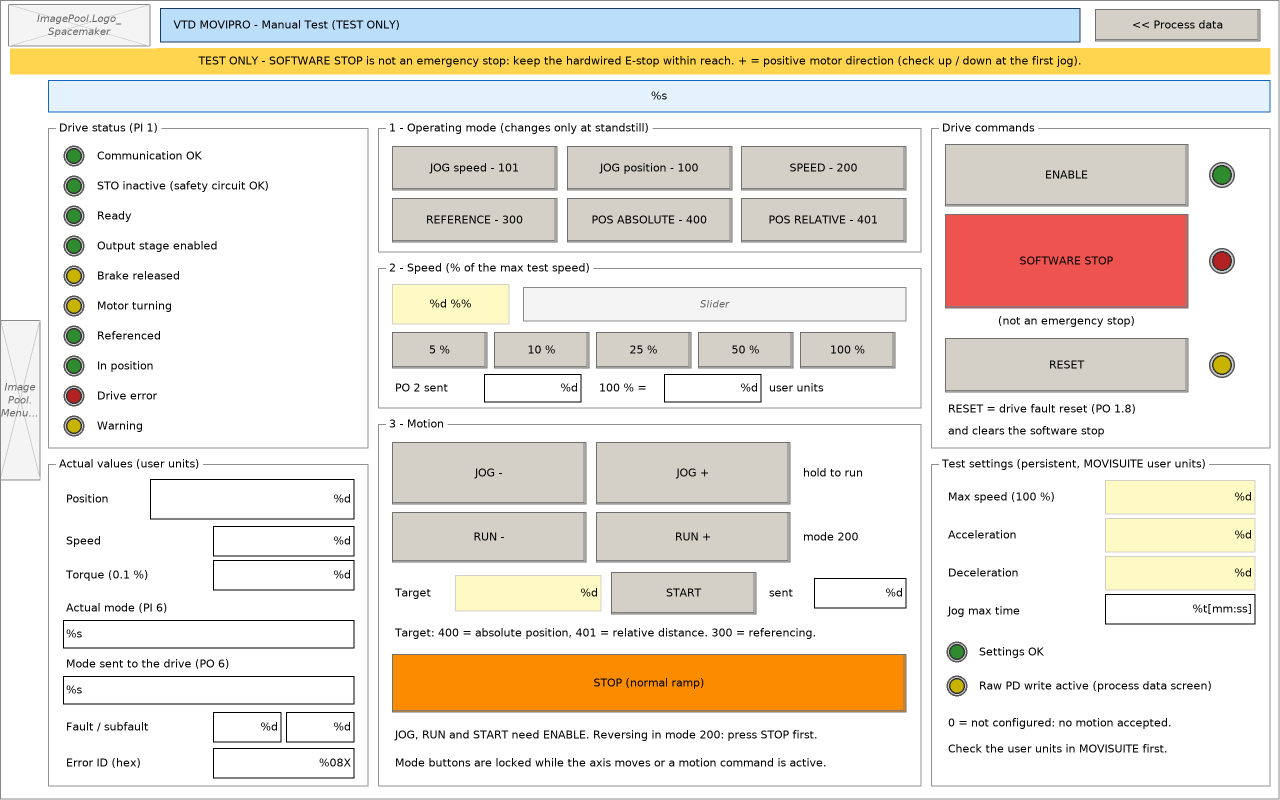
VISUALIZATION VTDManualTest  // 1280x800
    Rectangle (160,8 920x34), "VTD MOVIPRO - Manual Test (TEST ONLY)"
    Button (1095,9 165x32), "<< Process data"
        OnMouseClick: change screen: Visualization
    Rectangle (10,48 1260x26), "TEST ONLY - SOFTWARE STOP is not an emergency stop: keep the hardwired E-stop within reach. + = positive motor direction (check up / down at the first jog)."
    Rectangle (48,80 1222x32), "%s", text variable: GVL_HMI_VTD.stManualStatus.sMessage, colour toggle: GVL_HMI_VTD.stManualStatus.bMessageAlarm
    GroupBox (48,120 320x328), "Drive status (PI 1)"
    Lamp1 (62,144 24x24), variable: GVL_HMI_VTD.stManualStatus.stDrive.bCommunicationOk, style: Lamp-Lamp1-Green
    Rectangle (94,142 261x28), "Communication OK"
    Lamp1 (62,174 24x24), variable: GVL_HMI_VTD.stManualStatus.stDrive.bStoInactive, style: Lamp-Lamp1-Green
    Rectangle (94,172 261x28), "STO inactive (safety circuit OK)"
    Lamp1 (62,204 24x24), variable: GVL_HMI_VTD.stManualStatus.stDrive.bReady, style: Lamp-Lamp1-Green
    Rectangle (94,202 261x28), "Ready"
    Lamp1 (62,234 24x24), variable: GVL_HMI_VTD.stManualStatus.stDrive.bOutputStageEnabled, style: Lamp-Lamp1-Green
    Rectangle (94,232 261x28), "Output stage enabled"
    Lamp1 (62,264 24x24), variable: GVL_HMI_VTD.stManualStatus.stDrive.bBrakeReleased, style: Lamp-Lamp1-Yellow
    Rectangle (94,262 261x28), "Brake released"
    Lamp1 (62,294 24x24), variable: GVL_HMI_VTD.stManualStatus.stDrive.bMotorTurning, style: Lamp-Lamp1-Yellow
    Rectangle (94,292 261x28), "Motor turning"
    Lamp1 (62,324 24x24), variable: GVL_HMI_VTD.stManualStatus.stDrive.bReferenced, style: Lamp-Lamp1-Green
    Rectangle (94,322 261x28), "Referenced"
    Lamp1 (62,354 24x24), variable: GVL_HMI_VTD.stManualStatus.stDrive.bInPosition, style: Lamp-Lamp1-Green
    Rectangle (94,352 261x28), "In position"
    Lamp1 (62,384 24x24), variable: GVL_HMI_VTD.stManualStatus.stDrive.bError, style: Lamp-Lamp1-Red
    Rectangle (94,382 261x28), "Drive error"
    Lamp1 (62,414 24x24), variable: GVL_HMI_VTD.stManualStatus.stDrive.bWarning, style: Lamp-Lamp1-Yellow
    Rectangle (94,412 261x28), "Warning"
    GroupBox (48,456 320x330), "Actual values (user units)"
    Rectangle (63,484 82x30), "Position"
    Rectangle (150,479 204x40), "%d", text variable: GVL_HMI_VTD.stManualStatus.stDrive.diActualPosition
    Rectangle (63,526 145x30), "Speed"
    Rectangle (213,526 141x30), "%d", text variable: GVL_HMI_VTD.stManualStatus.stDrive.iActualSpeed
    Rectangle (63,560 145x30), "Torque (0.1 %)"
    Rectangle (213,560 141x30), "%d", text variable: GVL_HMI_VTD.stManualStatus.stDrive.iActualTorque_0p1pct
    Rectangle (63,596 291x24), "Actual mode (PI 6)"
    Rectangle (63,620 291x28), "%s", text variable: GVL_HMI_VTD.stManualStatus.sActualModeName
    Rectangle (63,652 291x24), "Mode sent to the drive (PO 6)"
    Rectangle (63,676 291x28), "%s", text variable: GVL_HMI_VTD.stManualStatus.sModeActiveName
    Rectangle (63,712 145x30), "Fault / subfault"
    Rectangle (213,712 68x30), "%d", text variable: GVL_HMI_VTD.stManualStatus.stDrive.byFaultCode
    Rectangle (286,712 68x30), "%d", text variable: GVL_HMI_VTD.stManualStatus.stDrive.bySubfaultCode
    Rectangle (63,748 145x30), "Error ID (hex)"
    Rectangle (213,748 141x30), "%08X", text variable: GVL_HMI_VTD.stManualStatus.udiErrorId
    GroupBox (378,120 543x132), "1 - Operating mode (changes only at standstill)"
    Button (392,146 165x44), "JOG speed - 101", colour toggle: GVL_HMI_VTD.stManualStatus.bModeJogSpeed, input disabled if: NOT GVL_HMI_VTD.stManualStatus.bModeChangeAllowed
        OnMouseClick: execute { GVL_HMI_VTD.stManualCommand.eModeRequest := E_SEW_MovikitMode.JogSpeedControlled; }
    Button (567,146 165x44), "JOG position - 100", colour toggle: GVL_HMI_VTD.stManualStatus.bModeJogPosition, input disabled if: NOT GVL_HMI_VTD.stManualStatus.bModeChangeAllowed
        OnMouseClick: execute { GVL_HMI_VTD.stManualCommand.eModeRequest := E_SEW_MovikitMode.JogPositionControlled; }
    Button (741,146 165x44), "SPEED - 200", colour toggle: GVL_HMI_VTD.stManualStatus.bModeSpeed, input disabled if: NOT GVL_HMI_VTD.stManualStatus.bModeChangeAllowed
        OnMouseClick: execute { GVL_HMI_VTD.stManualCommand.eModeRequest := E_SEW_MovikitMode.Speed; }
    Button (392,198 165x44), "REFERENCE - 300", colour toggle: GVL_HMI_VTD.stManualStatus.bModeReferencing, input disabled if: NOT GVL_HMI_VTD.stManualStatus.bModeChangeAllowed
        OnMouseClick: execute { GVL_HMI_VTD.stManualCommand.eModeRequest := E_SEW_MovikitMode.ReferencingOffsetConfigured; }
    Button (567,198 165x44), "POS ABSOLUTE - 400", colour toggle: GVL_HMI_VTD.stManualStatus.bModePositionAbsolute, input disabled if: NOT GVL_HMI_VTD.stManualStatus.bModeChangeAllowed
        OnMouseClick: execute { GVL_HMI_VTD.stManualCommand.eModeRequest := E_SEW_MovikitMode.PositioningAbsolute; }
    Button (741,198 165x44), "POS RELATIVE - 401", colour toggle: GVL_HMI_VTD.stManualStatus.bModePositionRelative, input disabled if: NOT GVL_HMI_VTD.stManualStatus.bModeChangeAllowed
        OnMouseClick: execute { GVL_HMI_VTD.stManualCommand.eModeRequest := E_SEW_MovikitMode.PositioningRelative; }
    GroupBox (378,260 543x148), "2 - Speed (% of the max test speed)"
    Textfield (392,284 117x40), "%d %%", text variable: GVL_HMI_VTD.stManualCommand.iSpeedPercent
        OnMouseClick: write the text variable via VisuDialogs.Numpad, min 0, max 100
    Slider (523,287 383x34), variable: GVL_HMI_VTD.stManualCommand.iSpeedPercent, scale 0..100
    Button (392,332 95x36), "5 %"
        OnMouseClick: execute { GVL_HMI_VTD.stManualCommand.iSpeedPercent := 5; }
    Button (494,332 95x36), "10 %"
        OnMouseClick: execute { GVL_HMI_VTD.stManualCommand.iSpeedPercent := 10; }
    Button (596,332 95x36), "25 %"
        OnMouseClick: execute { GVL_HMI_VTD.stManualCommand.iSpeedPercent := 25; }
    Button (698,332 95x36), "50 %"
        OnMouseClick: execute { GVL_HMI_VTD.stManualCommand.iSpeedPercent := 50; }
    Button (800,332 95x36), "100 %"
        OnMouseClick: execute { GVL_HMI_VTD.stManualCommand.iSpeedPercent := 100; }
    Rectangle (392,374 92x28), "PO 2 sent"
    Rectangle (484,374 97x28), "%d", text variable: GVL_HMI_VTD.stManualStatus.iSpeedSetpoint
    Rectangle (596,374 68x28), "100 % ="
    Rectangle (664,374 97x28), "%d", text variable: GVL_HMI_VTD.stManualSettings.iMaxSpeed
    Rectangle (766,374 140x28), "user units"
    GroupBox (378,416 543x370), "3 - Motion"
    Button (392,442 194x62), "JOG -", colour toggle: GVL_HMI_VTD.stManualStatus.bJogNegativeActive, input disabled if: NOT GVL_HMI_VTD.stManualStatus.bJogAvailable
        tap GVL_HMI_VTD.stManualCommand.bJogNegative p3779583253=TRUE
    Button (596,442 194x62), "JOG +", colour toggle: GVL_HMI_VTD.stManualStatus.bJogPositiveActive, input disabled if: NOT GVL_HMI_VTD.stManualStatus.bJogAvailable
        tap GVL_HMI_VTD.stManualCommand.bJogPositive p3779583253=TRUE
    Rectangle (800,458 111x30), "hold to run"
    Button (392,512 194x50), "RUN -", colour toggle: GVL_HMI_VTD.stManualStatus.bRunNegativeActive, input disabled if: NOT GVL_HMI_VTD.stManualStatus.bRunAvailable
        tap GVL_HMI_VTD.stManualCommand.bRunNegative p3779583253=TRUE
    Button (596,512 194x50), "RUN +", colour toggle: GVL_HMI_VTD.stManualStatus.bRunPositiveActive, input disabled if: NOT GVL_HMI_VTD.stManualStatus.bRunAvailable
        tap GVL_HMI_VTD.stManualCommand.bRunPositive p3779583253=TRUE
    Rectangle (800,522 111x30), "mode 200"
    Rectangle (392,578 63x30), "Target"
    Textfield (455,575 146x36), "%d", text variable: GVL_HMI_VTD.stManualCommand.diTargetPosition
        OnMouseClick: write the text variable via VisuDialogs.Numpad, min -2147483648, max 2147483647
    Button (611,572 145x42), "START", colour toggle: GVL_HMI_VTD.stManualStatus.bStartActive, input disabled if: NOT GVL_HMI_VTD.stManualStatus.bStartAvailable
        tap GVL_HMI_VTD.stManualCommand.bStart p3779583253=TRUE
    Rectangle (766,578 48x30), "sent"
    Rectangle (814,578 92x30), "%d", text variable: GVL_HMI_VTD.stManualStatus.diTargetPositionSent
    Rectangle (392,620 514x26), "Target: 400 = absolute position, 401 = relative distance. 300 = referencing."
    Button (392,654 514x58), "STOP (normal ramp)"
        tap GVL_HMI_VTD.stManualCommand.bStop p3779583253=TRUE
    Rectangle (392,722 514x26), "JOG, RUN and START need ENABLE. Reversing in mode 200: press STOP first."
    Rectangle (392,750 514x26), "Mode buttons are locked while the axis moves or a motion command is active."
    GroupBox (931,120 339x328), "Drive commands"
    Button (945,144 243x62), "ENABLE", colour toggle: GVL_HMI_VTD.stManualStatus.bEnableActive
        toggle GVL_HMI_VTD.stManualCommand.bEnable
    Lamp1 (1207,160 30x30), variable: GVL_HMI_VTD.stManualStatus.bEnableActive, style: Lamp-Lamp1-Green
    Button (945,214 243x94), "SOFTWARE STOP"
        tap GVL_HMI_VTD.stManualCommand.bSoftwareStop p3779583253=TRUE
    Lamp1 (1207,246 30x30), variable: GVL_HMI_VTD.stManualStatus.bSoftwareStopActive, style: Lamp-Lamp1-Red
    Rectangle (945,310 243x22), "(not an emergency stop)"
    Button (945,338 243x54), "RESET"
        tap GVL_HMI_VTD.stManualCommand.bReset p3779583253=TRUE
    Lamp1 (1207,350 30x30), variable: GVL_HMI_VTD.stManualStatus.bFaultResetActive, style: Lamp-Lamp1-Yellow
    Rectangle (945,398 315x22), "RESET = drive fault reset (PO 1.8)"
    Rectangle (945,420 315x22), "and clears the software stop"
    GroupBox (931,456 339x330), "Test settings (persistent, MOVISUITE user units)"
    Rectangle (945,482 155x30), "Max speed (100 %)"
    Textfield (1105,480 150x34), "%d", text variable: GVL_HMI_VTD.stManualSettings.iMaxSpeed
        OnMouseClick: write the text variable via VisuDialogs.Numpad, min 0, max 32767
    Rectangle (945,520 155x30), "Acceleration"
    Textfield (1105,518 150x34), "%d", text variable: GVL_HMI_VTD.stManualSettings.uiAcceleration
        OnMouseClick: write the text variable via VisuDialogs.Numpad, min 0, max 65535
    Rectangle (945,558 155x30), "Deceleration"
    Textfield (1105,556 150x34), "%d", text variable: GVL_HMI_VTD.stManualSettings.uiDeceleration
        OnMouseClick: write the text variable via VisuDialogs.Numpad, min 0, max 65535
    Rectangle (945,596 155x30), "Jog max time"
    Rectangle (1105,594 150x30), "%t[mm:ss]", text variable: GVL_HMI_VTD.stManualSettings.tJogMaxTime
    Lamp1 (945,640 24x24), variable: GVL_HMI_VTD.stManualStatus.bSettingsValid, style: Lamp-Lamp1-Green
    Rectangle (976,637 281x30), "Settings OK"
    Lamp1 (945,674 24x24), variable: GVL_HMI_VTD.stManualStatus.bRawWriteActive, style: Lamp-Lamp1-Yellow
    Rectangle (976,671 281x30), "Raw PD write active (process data screen)"
    Rectangle (945,710 315x26), "0 = not configured: no motion accepted."
    Rectangle (945,736 315x26), "Check the user units in MOVISUITE first."
    Rectangle (0,0 156x48)
        OnMouseClick: change screen: Main
    Image (8,4 142x42), image: ImagePool.Logo_Spacemaker
        OnMouseClick: change screen: Main
    Rectangle (0,320 40x160)
        OnMouseEnter: OpenDialog Dialog=Dialog, OpenModal=True, PositionX=0, PositionY=0
        OnMouseClick: OpenDialog Dialog=Dialog, OpenModal=True, PositionX=0, PositionY=0
    Image (0,320 40x160), image: ImagePool.Menu_Tab
        OnMouseEnter: OpenDialog Dialog=Dialog, OpenModal=True, PositionX=0, PositionY=0
        OnMouseClick: OpenDialog Dialog=Dialog, OpenModal=True, PositionX=0, PositionY=0
END_VISUALIZATION

(* stored: Version 1.1.0.1
   Visu VTDManualTest: Id {3c4ba5e1-66b9-42c1-b198-2293ecdc49e7} *)
